// TIA Portal V20 export
DATA_BLOCK "DataToSafety_DB"   // DB52
// stored: InstanceOfName DataToSafety, InstanceOfType FB
"DataToSafety"
   // VAR
   //    ACK_Taste : Bool := FALSE;
   //    BA_Manuell : Bool;
   //    BA_Automatik : Bool;
   //    BA_Verwaltung : Bool;
   //    BA_Richten : Bool;
   //    Ruekfuehrung_Bosch_Antriebe : Bool;
   // END_VAR
BEGIN
END_DATA_BLOCK
